{attribute 'qualified_only'}
{attribute 'strict'}
{attribute 'to_string'}
TYPE E_DWord :
(
	eOptionA := 0,
	eOptionB,
	eOptionC
) DWORD;
END_TYPE

(* stored: Version 1.1.0.1, ProductVersion 3.1.4026.19
   DUT E_DWord: Id {99bb4689-9462-4e19-aaa9-b766f1fe9a9f} *)
